// TIA Portal V21 export
// export: Created 2026-08-21T20:18:51.1003435Z, ExportSetting None, DisplayName Totally Integrated Automation Portal, DisplayVersion V21, DisplayName STEP 7 Professional, DisplayVersion V21, DisplayName STEP 7 Safety, DisplayVersion V21, DisplayName Tech WebApplication, DisplayVersion V21, DisplayName WinCC Basic/Comfort/Advanced, DisplayVersion V21, DisplayName WinCC Professional, DisplayVersion V21, DisplayName WinCC Unified, DisplayVersion V21
FUNCTION "FIT100_Liter" : Void   // FC15, FBD
{ S7_Optimized_Access := 'TRUE' }
// stored: SetENOAutomatically false
BEGIN

REGION Network 1: MonAnL
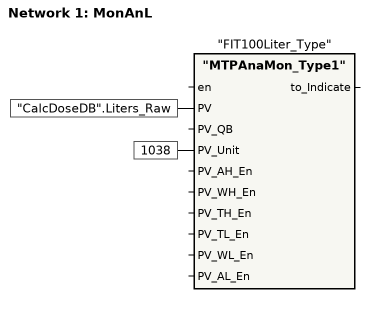
   "FIT100Liter_Type"(PV := "CalcDoseDB".Liters_Raw, PV_Unit := 1038);   // "MTPAnaMon_Type1"
END_REGION
END_FUNCTION
